{attribute 'pack_mode' := '1'}
TYPE ST_ProtectionConfigWirePacket :
STRUCT
	Header	:	ST_MqttCommandHeader;
	Record	:	ST_ProtectionConfig_Rx;	// DeviceIndex 없는 단일 레코드
END_STRUCT
END_TYPE

(* stored: Version 1.1.0.1, ProductVersion 3.1.4024.15
   DUT ST_ProtectionConfigWirePacket: Id {8c6d64ae-954f-499d-b545-17ff38b3cb87} *)
